(* IEC 61131-3 sources: nautilus/lang/conformance/fb-tof, 1 file *)

(* ---- fb-tof.st ---- *)
PROGRAM TofSt
(* TOF in Structured Text: the reference path. *)
VAR_EXTERNAL
    IN    : BOOL;
    PT    : TIME;
    st_Q  : BOOL;
    st_ET : TIME;
END_VAR
VAR
    t : TOF;
END_VAR

t(IN := IN, PT := PT);
st_Q  := t.Q;
st_ET := t.ET;
END_PROGRAM
